FUNCTION_BLOCK toffffblock
VAR_INPUT
	in:BOOL;
	pt:TIME;
END_VAR
VAR_OUTPUT
	out:BOOL;
	et:TIME;
END_VAR
VAR
	tstarttime:TIME;
	btiming:BOOL;
	bprevin:BOOL;
	
END_VAR

IF in THEN
	out:=TRUE;
	et:=T#0MS;
	btiming:=FALSE;
ELSE
	IF bprevin THEN
		tstarttime:=TIME();
		btiming:=TRUE;
		
		
	END_IF
	IF btiming THEN
		et:=TIME()-tstarttime;
		IF et>=pt THEN
			et:=pt;
			out:=FALSE;
			btiming:=FALSE;
			
		END_IF
	END_IF
END_IF
bprevin:=in;

END_FUNCTION_BLOCK

(* stored: Version 1.1.0.1, ProductVersion 3.1.4024.16
   POU toffffblock: Id {27e06b06-73a5-4efb-a636-6a6689930910}, SpecialFunc None *)
